// Mitsubishi GX Works2 project: 261012_타이머실습_타이머추가응용4   PLC: Q03UDV

PROGRAM MAIN
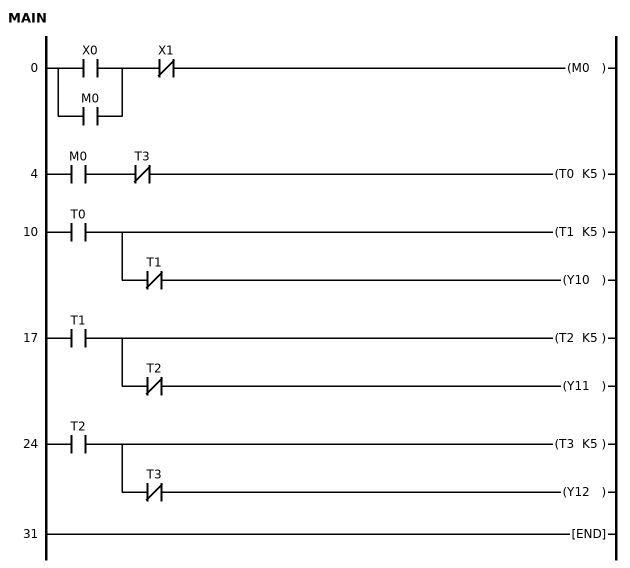
0     LD      X0
      OR      M0
      ANI     X1
      OUT     M0
4     LD      M0
      ANI     T3
      OUT     T0 K5
10    LD      T0
      OUT     T1 K5
      ANI     T1
      OUT     Y10
17    LD      T1
      OUT     T2 K5
      ANI     T2
      OUT     Y11
24    LD      T2
      OUT     T3 K5
      ANI     T3
      OUT     Y12
31    END
END_PROGRAM
